FUNCTION_BLOCK FB_Infeed
VAR_INPUT
END_VAR
VAR_OUTPUT
END_VAR
VAR
END_VAR

END_FUNCTION_BLOCK

(* stored: Version 1.1.0.1
   POU FB_Infeed: Id {e10d4917-c597-4ad2-a9c0-c75433bffb14}, SpecialFunc None *)
